Fanuc KAREL source: KD00073.KL

PROGRAM KD00073
%NOLOCKGROUP
VAR
  I: INTEGER
  J: INTEGER
  B: BOOLEAN
  R: REAL
  S: STRING[80]
BEGIN
  I = 0
  REPEAT
    I = I + 1
  UNTIL I > 2
END KD00073
